FUNCTION_BLOCK F (* Negative C2: two positions, but every scan goes through one common state and the position is forgotten there *)
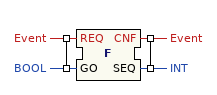
  EVENT_INPUT
    REQ WITH GO;
  END_EVENT
  EVENT_OUTPUT
    CNF WITH SEQ;
  END_EVENT
  VAR_INPUT
    GO : BOOL;
  END_VAR
  VAR_OUTPUT
    SEQ : INT;
  END_VAR
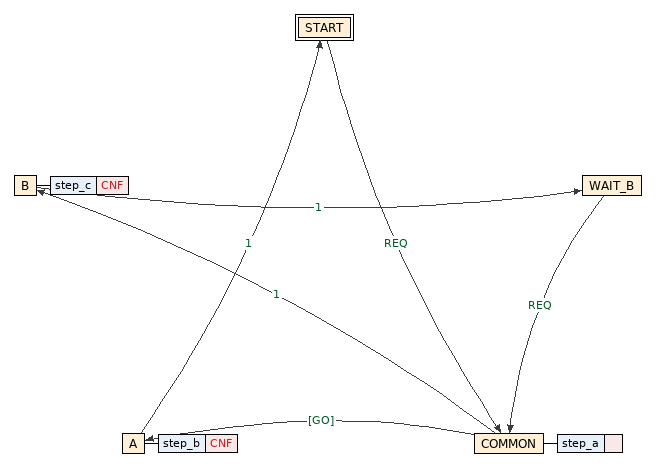
  EC_STATES
    START;
    WAIT_B;
    COMMON : step_a;
    A : step_b -> CNF;
    B : step_c -> CNF;
  END_STATES
  EC_TRANSITIONS
    START TO COMMON := REQ;
    WAIT_B TO COMMON := REQ;
    COMMON TO A := [GO];
    COMMON TO B := 1;
    A TO START := 1;
    B TO WAIT_B := 1;
  END_TRANSITIONS
  ALGORITHM step_a IN ST:
SEQ := 0;
IF GO THEN
  SEQ := 1;
END_IF;
  END_ALGORITHM
  ALGORITHM step_b IN ST:
IF NOT GO THEN
  SEQ := 0;
END_IF;
  END_ALGORITHM
  ALGORITHM step_c IN ST:
SEQ := 2;
  END_ALGORITHM
END_FUNCTION_BLOCK
